Fanuc KAREL source: KB00147.KL

PROGRAM KB00147
%NOLOCKGROUP
%ENVIRONMENT MEMO
VAR
  P1: STRING[80]
  P2: STRING[80]
  P3: STRING[80]
  P4: INTEGER
BEGIN
  P1 = 'A'
  P2 = 'A'
  P3 = 'A'
  P4 = 1
  RENAME_VAR(P1, P2, P3, P4)
END KB00147
